// TIA Portal V20 export
// export: Created 2026-10-19T18:45:52.4364559Z, ExportSetting None, DisplayName Totally Integrated Automation Portal, DisplayVersion V20 Update 6, DisplayName TIA Portal Openness, DisplayVersion V20 Update 6, DisplayName TIA Portal Version Control Interface, DisplayVersion V20 Update 6, DisplayName SINAMICS Startdrive Advanced, DisplayVersion V20 SP1, DisplayName SINAMICS Startdrive G130, G150, S120, S150, SINAMICS MV, G220, S200, S210, DisplayVersion V20 SP1, DisplayName SINAMICS Startdrive G110M, G120, G120C, G120D, G120P, G115D, DisplayVersion V20 SP1, DisplayName STEP 7 Professional, DisplayVersion V20 Update 6, DisplayName STEP 7 Safety, DisplayVersion V20 Update 2, DisplayName WinCC Basic/Comfort/Advanced, DisplayVersion V20 Update 6, DisplayName WinCC Unified, DisplayVersion V20 Update 6
VAR_GLOBAL   // PLC tag table "IO_Charger Panel_L5"
   "CHARGER L5 - Output Voltage" AT %ID848 : Real;   // Actual Output Voltage
   "CHARGER L5 - Output Current" AT %ID852 : Real;   // Actual Output Current
   "CHARGER L5 - Set Voltage Feedback" AT %ID856 : Real;   // Set Voltage Value
   "CHARGER L5 - Set Current Feedback" AT %ID860 : Real;   // Set Current Value
   "CHARGER L5 - Charging Start" AT %I864.0 : Bool;   // Charging Running Status
   "CHARGER L5 - Set Voltage Output" AT %QD424 : Real;   // Issue Target Voltage
   "CHARGER L5 - Set Current Output" AT %QD428 : Real;   // Issue Target Current
   "CHARGER L5 - Start Charging" AT %Q432.0 : Bool;   // Start Charging Command
   "CHARGER L5 - Stop Charging" AT %Q432.1 : Bool;   // Stop Charging Command
   "CHARGER L5 - Confirm Voltage & Current Setting" AT %Q432.2 : Bool;   // Confirmation Command
END_VAR
